Yaskawa INFORM job: MANYMOV.JBI

/JOB
//NAME MANYMOV
//POS
///NPOS 40,0,40,0,0,0
///TOOL 9
///POSTYPE PULSE
///PULSE
C00000=0,0,0
C00001=0,0,0
C00002=0,0,0
C00003=0,0,0
C00004=0,0,0
C00005=0,0,0
C00006=0,0,0
C00007=0,0,0
C00008=0,0,0
C00009=0,0,0
C00010=0,0,0
C00011=0,0,0
C00012=0,0,0
C00013=0,0,0
C00014=0,0,0
C00015=0,0,0
C00016=0,0,0
C00017=0,0,0
C00018=0,0,0
C00019=0,0,0
C00020=0,0,0
C00021=0,0,0
C00022=0,0,0
C00023=0,0,0
C00024=0,0,0
C00025=0,0,0
C00026=0,0,0
C00027=0,0,0
C00028=0,0,0
C00029=0,0,0
C00030=0,0,0
C00031=0,0,0
C00032=0,0,0
C00033=0,0,0
C00034=0,0,0
C00035=0,0,0
C00036=0,0,0
C00037=0,0,0
C00038=0,0,0
C00039=0,0,0
EC00000=0
EC00001=0
EC00002=0
EC00003=0
EC00004=0
EC00005=0
EC00006=0
EC00007=0
EC00008=0
EC00009=0
EC00010=0
EC00011=0
EC00012=0
EC00013=0
EC00014=0
EC00015=0
EC00016=0
EC00017=0
EC00018=0
EC00019=0
EC00020=0
EC00021=0
EC00022=0
EC00023=0
EC00024=0
EC00025=0
EC00026=0
EC00027=0
EC00028=0
EC00029=0
EC00030=0
EC00031=0
EC00032=0
EC00033=0
EC00034=0
EC00035=0
EC00036=0
EC00037=0
EC00038=0
EC00039=0
//INST
<volatile>
///COMM Generated using RoboDK
///ATTR SC,RW
///GROUP1 RB1
NOP
'Program generated by RoboDK v
'6.0.7 for Yaskawa Motoman EPL
'160 on XX/XX/XXXX 18:00:00
'Using nominal kinematics.
'Using Frame S (targets wrt ba
'se):
'1234.6,-98.8,50.5,0.0,0.0,30.
'0
'Tool Tool S should be close t
'o:
'10.0,20.0,150.0,0.0,0.0,0.0
MOVJ C00000 VJ=50.00  +MOVJ EC00000 VJ=100.00
MOVL C00001 V=500.0  +MOVJ EC00001 VJ=100.00
MOVJ C00002 VJ=50.00  +MOVJ EC00002 VJ=100.00
MOVL C00003 V=500.0  +MOVJ EC00003 VJ=100.00
MOVJ C00004 VJ=50.00  +MOVJ EC00004 VJ=100.00
MOVL C00005 V=500.0  +MOVJ EC00005 VJ=100.00
MOVJ C00006 VJ=50.00  +MOVJ EC00006 VJ=100.00
MOVL C00007 V=500.0  +MOVJ EC00007 VJ=100.00
MOVJ C00008 VJ=50.00  +MOVJ EC00008 VJ=100.00
MOVL C00009 V=500.0  +MOVJ EC00009 VJ=100.00
MOVJ C00010 VJ=50.00  +MOVJ EC00010 VJ=100.00
MOVL C00011 V=500.0  +MOVJ EC00011 VJ=100.00
MOVJ C00012 VJ=50.00  +MOVJ EC00012 VJ=100.00
MOVL C00013 V=500.0  +MOVJ EC00013 VJ=100.00
MOVJ C00014 VJ=50.00  +MOVJ EC00014 VJ=100.00
MOVL C00015 V=500.0  +MOVJ EC00015 VJ=100.00
MOVJ C00016 VJ=50.00  +MOVJ EC00016 VJ=100.00
MOVL C00017 V=500.0  +MOVJ EC00017 VJ=100.00
MOVJ C00018 VJ=50.00  +MOVJ EC00018 VJ=100.00
MOVL C00019 V=500.0  +MOVJ EC00019 VJ=100.00
MOVJ C00020 VJ=50.00  +MOVJ EC00020 VJ=100.00
MOVL C00021 V=500.0  +MOVJ EC00021 VJ=100.00
MOVJ C00022 VJ=50.00  +MOVJ EC00022 VJ=100.00
MOVL C00023 V=500.0  +MOVJ EC00023 VJ=100.00
MOVJ C00024 VJ=50.00  +MOVJ EC00024 VJ=100.00
MOVL C00025 V=500.0  +MOVJ EC00025 VJ=100.00
MOVJ C00026 VJ=50.00  +MOVJ EC00026 VJ=100.00
MOVL C00027 V=500.0  +MOVJ EC00027 VJ=100.00
MOVJ C00028 VJ=50.00  +MOVJ EC00028 VJ=100.00
MOVL C00029 V=500.0  +MOVJ EC00029 VJ=100.00
MOVJ C00030 VJ=50.00  +MOVJ EC00030 VJ=100.00
MOVL C00031 V=500.0  +MOVJ EC00031 VJ=100.00
MOVJ C00032 VJ=50.00  +MOVJ EC00032 VJ=100.00
MOVL C00033 V=500.0  +MOVJ EC00033 VJ=100.00
MOVJ C00034 VJ=50.00  +MOVJ EC00034 VJ=100.00
MOVL C00035 V=500.0  +MOVJ EC00035 VJ=100.00
MOVJ C00036 VJ=50.00  +MOVJ EC00036 VJ=100.00
MOVL C00037 V=500.0  +MOVJ EC00037 VJ=100.00
MOVJ C00038 VJ=50.00  +MOVJ EC00038 VJ=100.00
MOVL C00039 V=500.0  +MOVJ EC00039 VJ=100.00
END
